(* IEC 61131-3 sources: PLC_I/plc/src/cylinder, 18 files *)

(* ---- Cy确认.st ---- *)
(* 端位确认方式：传感器=真实信号连续有效，延时=动作后计时。 *)
TYPE Cy确认 :
(
    传感器 := 0,
    延时 := 1
);
END_TYPE

(* ---- Cy阀型.st ---- *)
(* 阀型枚举。数值顺序与协议类型一致，禁止插入或重排。 *)
TYPE Cy阀型 :
(
    单线圈复位 := 0,
    双线圈保持 := 1,
    真空吸附 := 2,
    真空带破真空 := 3
);
END_TYPE

(* ---- 结构体_Cy气缸配置.st ---- *)
(* 单缸配置：一行描述一个气缸的阀型、两侧绑定和确认方式。
   点地址是物理映像内的序号（输出 0..55，输入 0..111），不是 %QX/%IX 绝对地址。
   当前少量气缸全接内建点（直连模式）：点号 = 端子号（in动点 := 5 即 X5，
   out动点 := 2 即 Y2）；实际接线在 全局变量_物理IO.gvl.st 与
   程序_气缸输入映射/输出映射.st，本字段供 HMI 显示与配置校验。
   扩展模块缸点号从 32 起，由设备树映射到映像。
   选择 Cy确认.延时 时省略对应 in 字段；out原点 仅双线圈/真空带破真空使用。 *)
TYPE 结构体_Cy气缸配置 :
STRUCT
    已绑定 : BOOL;
    e阀型 : Cy阀型 := Cy阀型.单线圈复位;

    out动点 : WORD := 65535;
    out原点 : WORD := 65535;

    e动点确认 : Cy确认 := Cy确认.延时;
    in动点 : WORD := 65535;

    e原点确认 : Cy确认 := Cy确认.延时;
    in原点 : WORD := 65535;

    动点反相 : BOOL;
    原点反相 : BOOL;
END_STRUCT
END_TYPE

(* ---- 结构体_Cy状态.st ---- *)
(* 一次查询返回设备最近一次请求的状态，避免三个函数重复比对令牌。 *)
TYPE 结构体_Cy状态 :
STRUCT
    b忙 : BOOL;
    b完成 : BOOL;
    w故障 : WORD;
END_STRUCT
END_TYPE

(* ---- 结构体_Cy设备.st ---- *)
(* 设备运行态：保存最近一次业务请求号，业务代码不需要自己保存令牌。 *)
TYPE 结构体_Cy设备 :
STRUCT
    udi请求号 : UDINT;
    w错误 : WORD;
END_STRUCT
END_TYPE

(* ---- 结构体_气缸状态.st ---- *)
(* Volatile per-cylinder consumer state published for bound slots; zeros stay
   published for unbound cylinders. Written by PRG consumers after the Server. *)
TYPE 结构体_气缸状态 :
STRUCT
    b在动点 : BOOL;
    b在原点 : BOOL;
    b运动中 : BOOL;
    b故障 : BOOL;
    w错误码 : WORD;
END_STRUCT
END_TYPE

(* ---- 结构体_气缸请求.st ---- *)
TYPE 结构体_气缸请求 :
STRUCT
    udi请求号 : UDINT;
    udi完成号 : UDINT;
    w命令 : WORD;
    w错误 : WORD;
    b自动 : BOOL;
    b待下发 : BOOL;
    b忙 : BOOL;
END_STRUCT
END_TYPE

(* ---- 全局变量_Cy设备.gvl.st ---- *)
(* 设备编号：业务代码用名称表达设备，不用记数字。
   名称与现场绑定无关；未绑定设备调用动作会被拒绝。 *)
VAR_GLOBAL CONSTANT
    Cy夹紧 : UINT := 0;
    Cy定位 : UINT := 1;
END_VAR
VAR_GLOBAL
    (* 每个设备保存最近一次请求号，业务不需要自己管理令牌。 *)
    Cy设备状态 : ARRAY[0..53] OF 结构体_Cy设备;
END_VAR

(* ---- 全局变量_气缸请求.gvl.st ---- *)
{attribute 'qualified_only'}
VAR_GLOBAL
    ast请求 : ARRAY[0..53] OF 结构体_气缸请求;
    udi下个请求号 : UDINT;
    st许可快照 : 结构体_运行时;
END_VAR

(* ---- Cy动点.st ---- *)
(* 请求到动点/吸附。TRUE=已登记，内部保存请求号，业务无需自己持有。 *)
FUNCTION Cy动点 : BOOL
VAR_INPUT 设备 : UINT; END_VAR
Cy动点 := Cy提交(设备 := 设备, 命令 := 40);
END_FUNCTION

(* ---- Cy原点.st ---- *)
(* 请求到原点/释放。TRUE=已登记。 *)
FUNCTION Cy原点 : BOOL
VAR_INPUT 设备 : UINT; END_VAR
Cy原点 := Cy提交(设备 := 设备, 命令 := 41);
END_FUNCTION

(* ---- Cy取消.st ---- *)
(* 取消本次请求并撤销输出。TRUE=已登记；取消不代表到位。 *)
FUNCTION Cy取消 : BOOL
VAR_INPUT 设备 : UINT; END_VAR
Cy取消 := Cy提交(设备 := 设备, 命令 := 42);
END_FUNCTION

(* ---- Cy提交.st ---- *)
(* 业务语义API共用的请求号登记；拒绝时保留最近一次已接受请求。
   底层气缸_提交仍是所有来源唯一入槽/许可入口。 *)
FUNCTION Cy提交 : BOOL
VAR_INPUT
    设备 : UINT;
    命令 : WORD;
END_VAR
VAR
    udi请求号 : UDINT;
END_VAR
Cy提交 := FALSE;
IF 设备 >= 54 THEN RETURN; END_IF;
udi请求号 := 气缸_提交(缸号 := 设备, 命令 := 命令, 自动 := TRUE,
    Runtime := 全局变量_气缸请求.st许可快照);
IF udi请求号 = 0 THEN RETURN; END_IF;
Cy设备状态[设备].udi请求号 := udi请求号;
Cy提交 := TRUE;
END_FUNCTION

(* ---- Cy状态.st ---- *)
(* 设备最近一次请求的忙/完成/故障，令牌比对只在这里做一次。
   无请求返回故障 15；令牌失效（被其他来源替换）返回 19。 *)
FUNCTION Cy状态 : 结构体_Cy状态
VAR_INPUT 设备 : UINT; END_VAR
Cy状态.b忙 := FALSE;
Cy状态.b完成 := FALSE;
Cy状态.w故障 := ERR_非法;
IF 设备 >= 54 THEN
    RETURN;
END_IF;
IF Cy设备状态[设备].udi请求号 = 0 THEN
    RETURN;
END_IF;
Cy状态.w故障 := ERR_取消;
IF 全局变量_气缸请求.ast请求[设备].udi请求号 <> Cy设备状态[设备].udi请求号 THEN
    RETURN;
END_IF;
Cy状态.w故障 := 全局变量_气缸请求.ast请求[设备].w错误;
Cy状态.b忙 := 全局变量_气缸请求.ast请求[设备].b忙;
Cy状态.b完成 := (全局变量_气缸请求.ast请求[设备].udi完成号 = Cy设备状态[设备].udi请求号)
    AND NOT 全局变量_气缸请求.ast请求[设备].b忙;
END_FUNCTION

(* ---- 气缸_提交.st ---- *)
(* 所有来源唯一单槽入口。返回0拒绝，否则返回调用者必须保存的请求号。 *)
FUNCTION 气缸_提交 : UDINT
VAR_INPUT
    缸号 : UINT;
    命令 : WORD;
    自动 : BOOL;
END_VAR
VAR_IN_OUT
    Runtime : 结构体_运行时;
END_VAR
VAR
    w许可 : WORD;
END_VAR
气缸_提交 := 0;
IF 缸号 >= 54 THEN RETURN; END_IF;
IF (命令 <> 40) AND (命令 <> 41) AND (命令 <> 42) THEN RETURN; END_IF;
w许可 := 函数_动作许可(Code := 命令, ObjectWord := WORD#16#0200 OR UINT_TO_WORD(缸号),
    HmiOnline := Runtime.bHMI在线, JogBusy := FALSE, Resetting := Runtime.b复位中,
    b自动请求 := 自动, Runtime := Runtime, Store := 全局变量_保持区.Store);
IF w许可 <> 0 THEN RETURN; END_IF;
(* 42可覆盖任何请求；普通动作不能覆盖忙或尚未消费的停止。 *)
IF (命令 <> 42) AND (全局变量_气缸请求.ast请求[缸号].b忙
    OR 全局变量_气缸请求.ast请求[缸号].b待下发) THEN RETURN; END_IF;
IF 全局变量_气缸请求.udi下个请求号 = UDINT#4294967295 THEN
    全局变量_气缸请求.udi下个请求号 := 1;
ELSE
    全局变量_气缸请求.udi下个请求号 := 全局变量_气缸请求.udi下个请求号 + 1;
END_IF;
全局变量_气缸请求.ast请求[缸号].udi请求号 := 全局变量_气缸请求.udi下个请求号;
全局变量_气缸请求.ast请求[缸号].udi完成号 := 0;
全局变量_气缸请求.ast请求[缸号].w命令 := 命令;
全局变量_气缸请求.ast请求[缸号].w错误 := 0;
全局变量_气缸请求.ast请求[缸号].b自动 := 自动;
全局变量_气缸请求.ast请求[缸号].b待下发 := TRUE;
全局变量_气缸请求.ast请求[缸号].b忙 := TRUE;
气缸_提交 := 全局变量_气缸请求.udi下个请求号;
END_FUNCTION

(* ---- 气缸_配置有效.st ---- *)
FUNCTION 气缸_配置有效 : BOOL
VAR_INPUT 缸号 : UINT; END_VAR
VAR_IN_OUT Store : 结构体_配置; END_VAR
VAR i : UINT; j : UINT; k : UINT; w类型 : WORD; END_VAR
气缸_配置有效 := FALSE;
IF 缸号 >= 54 THEN RETURN; END_IF;
IF (Store.aw气缸配置[缸号, 0] AND WORD#16#FFF0) <> 0 THEN RETURN; END_IF;
w类型 := Store.aw气缸配置[缸号, 0] AND 3;
(* 输出地址按输出映像容量校验，输入地址按输入映像容量校验。 *)
FOR i := 1 TO 2 DO
    IF (Store.aw气缸配置[缸号, i] <> WORD#16#FFFF) AND (WORD_TO_UINT(Store.aw气缸配置[缸号, i]) >= ui气缸输出点数) THEN RETURN; END_IF;
END_FOR;
FOR i := 3 TO 4 DO
    IF (Store.aw气缸配置[缸号, i] <> WORD#16#FFFF) AND (WORD_TO_UINT(Store.aw气缸配置[缸号, i]) >= ui气缸输入点数) THEN RETURN; END_IF;
END_FOR;
IF Store.aw气缸配置[缸号, 1] = WORD#16#FFFF THEN RETURN; END_IF;
IF (w类型 = 0) OR (w类型 = 2) THEN
    IF Store.aw气缸配置[缸号, 2] <> WORD#16#FFFF THEN RETURN; END_IF;
ELSE
    IF (Store.aw气缸配置[缸号, 2] = WORD#16#FFFF)
        OR (Store.aw气缸配置[缸号, 2] = Store.aw气缸配置[缸号, 1]) THEN RETURN; END_IF;
END_IF;
IF (Store.aw气缸配置[缸号, 6] = 0)
    OR (Store.aw气缸配置[缸号, 5] >= Store.aw气缸配置[缸号, 6])
    OR (Store.aw气缸配置[缸号, 7] >= Store.aw气缸配置[缸号, 6]) THEN RETURN; END_IF;
IF ((Store.aw气缸配置[缸号, 3] = WORD#16#FFFF) AND (Store.aw气缸配置[缸号, 5] = 0))
    OR ((Store.aw气缸配置[缸号, 4] = WORD#16#FFFF) AND (Store.aw气缸配置[缸号, 7] = 0)) THEN RETURN; END_IF;
IF (Store.aw气缸配置[缸号, 3] <> WORD#16#FFFF)
    AND (Store.aw气缸配置[缸号, 3] = Store.aw气缸配置[缸号, 4]) THEN RETURN; END_IF;
(* 同一物理地址只能属于一个已绑定气缸：输出和输入都查重，
   防止两个缸抢同一个阀或同一个端位传感器。 *)
FOR i := 0 TO 53 DO
    IF (i <> 缸号) AND ((lw已绑定气缸 AND SHL(LWORD#1, i)) <> 0) THEN
        (* DI与DO是独立地址空间：仅在同类映像内查重。 *)
        FOR j := 1 TO 2 DO
            FOR k := 1 TO 2 DO
                IF (Store.aw气缸配置[缸号, j] <> WORD#16#FFFF)
                    AND (Store.aw气缸配置[缸号, j] = Store.aw气缸配置[i, k]) THEN RETURN; END_IF;
            END_FOR;
        END_FOR;
        FOR j := 3 TO 4 DO
            FOR k := 3 TO 4 DO
                IF (Store.aw气缸配置[缸号, j] <> WORD#16#FFFF)
                    AND (Store.aw气缸配置[缸号, j] = Store.aw气缸配置[i, k]) THEN RETURN; END_IF;
            END_FOR;
        END_FOR;
    END_IF;
END_FOR;
气缸_配置有效 := TRUE;
END_FUNCTION

(* ---- 功能块_气缸.st ---- *)
(* 单任务调用。输入为真实传感器，经调用者按存在性与极性归一。
   Token是内部UDINT请求号；连续扫描Execute=TRUE的新Token也可靠受理。
   CancelMode=1撤销完成资格并保持夹持输出（类型3关闭破真空），2撤销全部输出。
   本软件不是物理安全回路。 *)
FUNCTION_BLOCK 功能块_气缸
VAR_INPUT
    Execute : BOOL;
    Token : UDINT;
    Code : WORD;
    SensorWork : BOOL;
    SensorOrigin : BOOL;
    HasWorkSensor : BOOL := TRUE;
    HasOriginSensor : BOOL := TRUE;
    DelayMs : WORD;
    HomeDelayMs : WORD;
    TimeoutMs : WORD;
    HardEstop : BOOL;
    CancelMode : BYTE;
    ValveType : BYTE;
END_VAR
VAR_OUTPUT
    WorkOutput : BOOL;
    OriginOutput : BOOL;
    Moving : BOOL;
    Fault : BOOL;
    AtWork : BOOL;
    AtOrigin : BOOL;
    Error : WORD;
    DoneToken : UDINT;
END_VAR
VAR
    tmr动点滤波 : TON;
    tmr原点滤波 : TON;
    tmr运动 : TON;
    udi上次请求 : UDINT;
    udi活动请求 : UDINT;
    b新请求 : BOOL;
    b配置有效 : BOOL;
    b冲突 : BOOL;
    b取消 : BOOL;
    i目标侧 : INT;
    by锁定阀型 : BYTE;
    w锁定动点延时 : WORD;
    w锁定原点延时 : WORD;
    w锁定超时 : WORD;
    b锁定动点传感器 : BOOL;
    b锁定原点传感器 : BOOL;
END_VAR
b新请求 := Execute AND (Token <> 0) AND (Token <> udi上次请求);
IF b新请求 THEN udi上次请求 := Token; END_IF;
b配置有效 := (TimeoutMs > 0) AND (DelayMs < TimeoutMs) AND (HomeDelayMs < TimeoutMs)
    AND (ValveType <= 3) AND (HasWorkSensor OR (DelayMs > 0))
    AND (HasOriginSensor OR (HomeDelayMs > 0));
b冲突 := HasWorkSensor AND HasOriginSensor AND SensorWork AND SensorOrigin;
IF b新请求 AND (Code = 42) AND NOT HardEstop AND b配置有效 AND NOT b冲突 THEN
    Fault := FALSE; Error := 0;
END_IF;
IF HardEstop THEN Fault := TRUE; Error := 2103;
ELSIF NOT b配置有效 THEN Fault := TRUE; Error := 2131;
ELSIF b冲突 THEN Fault := TRUE; Error := 2110;
ELSIF (udi活动请求 <> 0) AND (DoneToken = 0) AND NOT (b新请求 AND (Code = 42))
    AND ((ValveType <> by锁定阀型)
    OR (DelayMs <> w锁定动点延时) OR (HomeDelayMs <> w锁定原点延时)
    OR (TimeoutMs <> w锁定超时) OR (HasWorkSensor <> b锁定动点传感器)
    OR (HasOriginSensor <> b锁定原点传感器)) THEN
    Fault := TRUE; Error := 2131;
END_IF;
b取消 := HardEstop OR Fault OR (CancelMode <> 0) OR (b新请求 AND (Code = 42));
IF b取消 THEN
    udi活动请求 := 0; DoneToken := 0; i目标侧 := 0; Moving := FALSE;
    IF HardEstop OR (CancelMode = 2) OR (b新请求 AND (Code = 42)) THEN
        WorkOutput := FALSE; OriginOutput := FALSE;
    ELSIF Fault THEN
        (* 真空只保持现有吸附；破真空必须关闭，等待人工42确认。 *)
        IF (ValveType <> 2) AND (ValveType <> 3) THEN
            WorkOutput := FALSE; OriginOutput := FALSE;
        ELSIF ValveType = 3 THEN
            OriginOutput := FALSE;
        END_IF;
    ELSIF ValveType = 3 THEN
        OriginOutput := FALSE;
    END_IF;
ELSIF b新请求 AND ((Code = 40) OR (Code = 41)) THEN
    udi活动请求 := Token; DoneToken := 0;
    IF Code = 40 THEN i目标侧 := 1; ELSE i目标侧 := 2; END_IF;
    by锁定阀型 := ValveType;
    w锁定动点延时 := DelayMs; w锁定原点延时 := HomeDelayMs; w锁定超时 := TimeoutMs;
    b锁定动点传感器 := HasWorkSensor; b锁定原点传感器 := HasOriginSensor;
    WorkOutput := i目标侧 = 1;
    OriginOutput := (i目标侧 = 2) AND ((ValveType = 1) OR (ValveType = 3));
END_IF;
(* 重置定时器后，同一扫描即开始新请求计时，包括单线圈无输出的回原动作。 *)
IF b新请求 OR b取消 THEN
    tmr动点滤波(IN := FALSE, PT := WORD_TO_TIME(DelayMs));
    tmr原点滤波(IN := FALSE, PT := WORD_TO_TIME(HomeDelayMs));
    tmr运动(IN := FALSE, PT := WORD_TO_TIME(TimeoutMs));
END_IF;
tmr动点滤波(IN := NOT b取消 AND ((HasWorkSensor AND SensorWork)
    OR (NOT HasWorkSensor AND (i目标侧 = 1) AND (udi活动请求 <> 0))), PT := WORD_TO_TIME(DelayMs));
tmr原点滤波(IN := NOT b取消 AND ((HasOriginSensor AND SensorOrigin)
    OR (NOT HasOriginSensor AND (i目标侧 = 2) AND (udi活动请求 <> 0))), PT := WORD_TO_TIME(HomeDelayMs));
AtWork := NOT b取消 AND tmr动点滤波.Q AND (NOT HasWorkSensor OR SensorWork);
AtOrigin := NOT b取消 AND tmr原点滤波.Q AND (NOT HasOriginSensor OR SensorOrigin);
(* 无感完成是本次请求的锁存估算，完成后修改延时不能使其闪断。 *)
IF NOT b取消 AND (DoneToken <> 0) THEN
    IF NOT HasWorkSensor THEN AtWork := i目标侧 = 1; END_IF;
    IF NOT HasOriginSensor THEN AtOrigin := i目标侧 = 2; END_IF;
END_IF;
Moving := NOT b取消 AND (udi活动请求 <> 0) AND (DoneToken = 0);
(* 总超时覆盖整个动作；同时到期时超时优先。 *)
tmr运动(IN := Moving, PT := WORD_TO_TIME(TimeoutMs));
IF tmr运动.Q THEN
    Fault := TRUE; Error := 2140; DoneToken := 0; udi活动请求 := 0; i目标侧 := 0;
    Moving := FALSE; AtWork := FALSE; AtOrigin := FALSE;
    (* 超时只保持现有吸附；类型3的破真空不得持续通电。 *)
    IF (ValveType <> 2) AND (ValveType <> 3) THEN
        WorkOutput := FALSE; OriginOutput := FALSE;
    ELSIF ValveType = 3 THEN
        OriginOutput := FALSE;
    END_IF;
ELSIF Moving AND (((i目标侧 = 1) AND AtWork) OR ((i目标侧 = 2) AND AtOrigin)) THEN
    DoneToken := udi活动请求; Moving := FALSE;
    IF (ValveType = 3) AND (i目标侧 = 2) THEN OriginOutput := FALSE; END_IF;
END_IF;
END_FUNCTION_BLOCK

(* ---- 功能块_气缸调度.st ---- *)
(* 唯一消费者：在服务端及本扫描模式更新之后运行。 *)
FUNCTION_BLOCK 功能块_气缸调度
VAR_INPUT StopAll : BOOL; END_VAR
VAR_IN_OUT Runtime : 结构体_运行时; END_VAR
VAR
    afb驱动 : ARRAY[0..53] OF 功能块_气缸;
    i : UINT;
    by取消 : BYTE;
    w许可 : WORD;
    b执行 : BOOL;
    b绑定 : BOOL;
    b动点传感器 : BOOL;
    b原点传感器 : BOOL;
END_VAR
FOR i := 0 TO 53 DO
    b绑定 := (lw已绑定气缸 AND SHL(LWORD#1, i)) <> 0;
    by取消 := 0;
    IF Runtime.b暂停 THEN by取消 := 1; END_IF;
    IF NOT Runtime.bHMI在线 OR Runtime.b复位中
        OR (全局变量_气缸请求.ast请求[i].b自动 AND (Runtime.b待复位 OR NOT Runtime.b运行 OR Runtime.b手动))
        OR (NOT 全局变量_气缸请求.ast请求[i].b自动 AND NOT Runtime.b手动) THEN
        by取消 := 1;
    END_IF;
    IF StopAll OR NOT b绑定 OR NOT ab气缸映射有效[i] OR NOT ab气缸模块就绪[i]
        OR Runtime.b硬急停 OR Runtime.b软急停 THEN by取消 := 2; END_IF;
    b执行 := 全局变量_气缸请求.ast请求[i].b待下发;
    (* 停止不受模式取消阻挡，始终能撤销输出并确认已消失的故障。 *)
    IF b执行 AND (全局变量_气缸请求.ast请求[i].w命令 <> 42) THEN
        w许可 := 函数_动作许可(Code := 全局变量_气缸请求.ast请求[i].w命令,
            ObjectWord := WORD#16#0200 OR UINT_TO_WORD(i), HmiOnline := Runtime.bHMI在线,
            JogBusy := FALSE, Resetting := Runtime.b复位中,
            b自动请求 := 全局变量_气缸请求.ast请求[i].b自动, b气缸已受理 := TRUE,
            Runtime := Runtime, Store := 全局变量_保持区.Store);
        IF w许可 <> 0 THEN
            b执行 := FALSE;
            全局变量_气缸请求.ast请求[i].w错误 := w许可;
            IF by取消 = 0 THEN by取消 := 1; END_IF;
        END_IF;
    END_IF;
    b动点传感器 := 全局变量_保持区.Store.aw气缸配置[i, 3] <> WORD#16#FFFF;
    b原点传感器 := 全局变量_保持区.Store.aw气缸配置[i, 4] <> WORD#16#FFFF;
    afb驱动[i](Execute := b执行, Token := 全局变量_气缸请求.ast请求[i].udi请求号,
        Code := 全局变量_气缸请求.ast请求[i].w命令,
        SensorWork := b动点传感器 AND (ab气缸动点传感器[i] XOR ((全局变量_保持区.Store.aw气缸配置[i, 0] AND 4) <> 0)),
        SensorOrigin := b原点传感器 AND (ab气缸原点传感器[i] XOR ((全局变量_保持区.Store.aw气缸配置[i, 0] AND 8) <> 0)),
        HasWorkSensor := b动点传感器, HasOriginSensor := b原点传感器,
        DelayMs := 全局变量_保持区.Store.aw气缸配置[i, 5], HomeDelayMs := 全局变量_保持区.Store.aw气缸配置[i, 7],
        TimeoutMs := 全局变量_保持区.Store.aw气缸配置[i, 6],
        ValveType := WORD_TO_BYTE(全局变量_保持区.Store.aw气缸配置[i, 0] AND 3),
        HardEstop := Runtime.b硬急停 OR Runtime.b软急停, CancelMode := by取消);
    全局变量_气缸请求.ast请求[i].b待下发 := FALSE;
    IF (by取消 <> 0) OR afb驱动[i].Fault OR (b执行 AND (全局变量_气缸请求.ast请求[i].w命令 = 42)) THEN
        全局变量_气缸请求.ast请求[i].b忙 := FALSE;
        全局变量_气缸请求.ast请求[i].udi完成号 := 0;
        IF afb驱动[i].Fault THEN 全局变量_气缸请求.ast请求[i].w错误 := afb驱动[i].Error;
        ELSIF 全局变量_气缸请求.ast请求[i].w错误 = 0 THEN 全局变量_气缸请求.ast请求[i].w错误 := 19;
        END_IF;
    ELSIF (afb驱动[i].DoneToken <> 0) AND (afb驱动[i].DoneToken = 全局变量_气缸请求.ast请求[i].udi请求号) THEN
        全局变量_气缸请求.ast请求[i].udi完成号 := afb驱动[i].DoneToken;
        全局变量_气缸请求.ast请求[i].b忙 := FALSE;
    END_IF;
    Runtime.ast气缸[i].b在动点 := afb驱动[i].AtWork;
    Runtime.ast气缸[i].b在原点 := afb驱动[i].AtOrigin;
    Runtime.ast气缸[i].b运动中 := afb驱动[i].Moving;
    Runtime.ast气缸[i].b故障 := afb驱动[i].Fault;
    Runtime.ast气缸[i].w错误码 := afb驱动[i].Error;
    ab气缸动点输出[i] := b绑定 AND ab气缸映射有效[i] AND ab气缸模块就绪[i] AND afb驱动[i].WorkOutput;
    ab气缸原点输出[i] := b绑定 AND ab气缸映射有效[i] AND ab气缸模块就绪[i] AND afb驱动[i].OriginOutput;
END_FOR;
全局变量_气缸请求.st许可快照 := Runtime;
END_FUNCTION_BLOCK
